TYPE ST_MotorStatus :
STRUCT
    //------------------------------------------------------------------
    // State machine
    //------------------------------------------------------------------
    eState              : E_MotorState;
    eControlMode        : E_ControlMode;

    //------------------------------------------------------------------
    // Status flags
    //------------------------------------------------------------------
    bEnabled            : BOOL;     // Drive power is on and ready
    bMoving             : BOOL;     // Axis is in motion
    bAtTarget           : BOOL;     // Position/velocity within tolerance
    bHomingDone         : BOOL;     // Homing completed successfully
    bZeroDone           : BOOL;     // Zero position completed successfully
    bTorqueActive       : BOOL;     // Torque control is active
    bTorqueInTorque     : BOOL;     // Target torque reached
    bError              : BOOL;     // Fault active
    nErrorID            : UDINT;    // TwinCAT NC error code (0 = no error)
    nResetStage         : BYTE;     // fault-recovery progress: 0 idle | 1 SoE drive
                                    // reset | 2 settle | 3 NC reset

    //------------------------------------------------------------------
    // Actual values
    //------------------------------------------------------------------
    fActPosition        : LREAL;    // [units]
    fActVelocity        : LREAL;    // [units/s]
    fActTorque          : LREAL;    // [% of rated torque]

    //------------------------------------------------------------------
    // Diagnostics
    //------------------------------------------------------------------
    fDcBusVoltage       : LREAL;    // [V]  — requires drive PDO mapping
    fDriveTemp          : LREAL;    // [°C] — requires drive PDO mapping
    nTimestamp          : UDINT;    // [ms since PLC start]
END_STRUCT
END_TYPE

(* stored: Version 1.1.0.1, ProductVersion 3.1.4026.18
   DUT ST_MotorStatus: Id {1d9fb2bb-4bf7-4960-a2c5-73a6bb6bc4c9} *)
